// TIA Portal V19 export
// export: Created 2026-10-15T09:44:22.91914Z, ExportSetting WithDefaults, DisplayName Totally Integrated Automation Portal, DisplayVersion V19, DisplayName TIA Portal Openness, DisplayVersion V19, DisplayName TIA Portal Version Control Interface, DisplayVersion V19, DisplayName STEP 7 Professional, DisplayVersion V19, DisplayName STEP 7 Safety, DisplayVersion V19, DisplayName WinCC Basic/Comfort/Advanced, DisplayVersion V19, DisplayName WinCC Unified, DisplayVersion V19
FUNCTION "ROLL_SetMWord" : Void   // FC2, SCL
{ S7_Optimized_Access := 'TRUE' }
VERSION : 0.1
// stored: AutoNumber true, IsIECCheckEnabled false, SetENOAutomatically false, UDAEnableTagReadback false
   VAR_INPUT
      FirstByte : Int;
      Value : Word;
   END_VAR
   VAR_TEMP
      bit : Int;
   END_VAR
BEGIN

   IF (#FirstByte < 0) OR (#FirstByte > 254) THEN
       "ROLL_IO".ConversionFault := TRUE;
       RETURN;
   END_IF;
   FOR #bit := 0 TO 7 DO
       "ROLL_State".M[#FirstByte, #bit] := (#Value AND SHL(IN := W#16#0001, N := #bit + 8)) <> W#16#0000;
       "ROLL_State".M[#FirstByte + 1, #bit] := (#Value AND SHL(IN := W#16#0001, N := #bit)) <> W#16#0000;
   END_FOR;
END_FUNCTION
